(*
SPDX-FileCopyrightText: c 2026 Oleksandr Tiutyk <trofimich@gmail.com>
SPDX-License-Identifier: MIT
License: https://opensource.org/license/mit
*)

(*!
<summary>Checks borrowed replacement and the surrounding entries.</summary>
<description>
Borrows a group-owned list reserved for this case. Use from one task at a stable address.
Teardown clears the list before publication.
</description>
*)

{attribute 'no_assign'}
{attribute 'no_explicit_call' := 'do not call this function block directly'}
FUNCTION_BLOCK ListGetAndSetGenericTest EXTENDS TOF_Testing.SingleCycleTest
VAR_STAT
	{attribute 'hide'}
	_ClassName : STRING := __POUNAME();
END_VAR
VAR
	_List : TOF_Collections.IList;
	_Values : ARRAY [0..5] OF STRING := ['String0', 'String1', 'String2', 'String3', 'String4', 'String5'];
END_VAR

(*!
<summary>Clears the fixture before the runner publishes the result.</summary>
<description>
Also runs after an unexpected exception interrupts the case.
</description>
*)
METHOD PROTECTED AfterTest
_List.Clear();
END_METHOD

//! <summary>Borrows the concrete class name. Callers must not modify it.</summary>
{attribute 'monitoring' := 'call'}
PROPERTY ClassName : REFERENCE TO STRING
GET
ClassName REF= _ClassName;
END_GET
END_PROPERTY

(*!
<summary>Checks borrowed replacement and the surrounding entries.</summary>
*)
METHOD PROTECTED ExecuteTest
VAR
	values : ARRAY [0..5] OF STRING := ['String0', 'String1', 'String2', 'String3', 'String4', 'String5'];
	entry : TOF_Core.GENERIC_VALUE;
	expected : ARRAY [0..2] OF STRING := ['String0', 'String4', 'String2'];
	i : DINT;
END_VAR
_List.AppendCopy(value := values[0]);
_List.AppendCopy(value := values[1]);
_List.AppendCopy(value := values[2]);

entry := TOF_Core.GenericValueFactory.FromStringReference(value := _Values[4]);
_List.SetGeneric(index := 1, value := entry);

Assert.ThatBool(
	actual := _List.Get(index := 1).Address = entry.Address AND_THEN NOT _List.Get(index := 1).IsMemoryOwner,
	message := "SetGeneric must retain the borrowed address and ownership mode"
).IsTrue();

Assert.ThatDInt(
	actual := _List.Length,
	message := "Unexpected sequence after GetAndSetGeneric length"
).ToBe(expected := DINT#3);

FOR i := 0 TO 2 DO
	Assert.ThatString(
		actual := _List.Get(index := i).AsString255(),
		message := TOF_Core.WideStrings.Concat255("Unexpected sequence after GetAndSetGeneric at index ", TO_WSTRING(i))
	).ToBe(expected := expected[i]);
END_FOR
END_METHOD

(*!
<summary>Binds the list fixture for this case.</summary>
<description>
Stores a borrowed interface without invoking the fixture. The owning group keeps it alive and
reserves it for this case. TestElement initializes the name and parent.
</description>
<param name="name">Display name of this case.</param>
<param name="parent">Group that owns this case.</param>
<param name="list">Required live list reserved for this case.</param>
*)
METHOD FB_init : BOOL
VAR_INPUT
	bInitRetains: BOOL; // TRUE: the retain variables are initialized (reset warm / reset cold)
	bInCopyCode: BOOL; // TRUE: the instance will be copied to the copy code afterward (online change)
	name : WSTRING;
	parent : TOF_Testing.ITestElement;
	list : TOF_Collections.IList;
END_VAR
_List := list;
FB_init := TRUE;
END_METHOD

//! <summary>Borrows the compiler-initialized namespace name. Callers must not modify it.</summary>
{attribute 'monitoring' := 'call'}
PROPERTY NamespaceName : REFERENCE TO STRING
GET
NamespaceName REF= CurrentNamespace.Name;
END_GET
END_PROPERTY

//! <summary>Reports the concrete instance size in bytes.</summary>
{attribute 'monitoring' := 'call'}
PROPERTY SelfSize : ULINT
GET
SelfSize := XSIZEOF(THIS^);
END_GET
END_PROPERTY

END_FUNCTION_BLOCK

(* stored: Version 1.1.0.1, ProductVersion 3.1.4026.21
   POU ListGetAndSetGenericTest: Id {d176b575-9771-488c-8b31-096adaf3f0a5}, SpecialFunc None
   Method AfterTest: Id {47dab618-db6d-4193-86b8-e47639b1c8b2}
   Property ClassName: Id {719f5628-a35e-4142-b59c-932d32472736}
   Get Get: Id {8edcaff4-35f6-4afe-bcbf-94bbc697c353}
   Method ExecuteTest: Id {f8163c98-a957-4f36-833c-6872db4476dd}
   Method FB_init: Id {c46b30f2-3e9d-40a3-bfcb-cac1da134a49}
   Property NamespaceName: Id {7bcb5d87-a577-40fa-87b8-c05a32cb1870}
   Get Get: Id {76a87593-316f-4c91-96c5-3ecb6cb89d3a}
   Property SelfSize: Id {2907363d-36e9-4e57-b238-a3d8a567b0fb}
   Get Get: Id {e5046cb5-b1f3-4df6-b15e-bc7f7b33176e} *)
